(* IEC 61131-3 sources: AyCD/codesys/src/POUs, 8 files *)

(* ---- COM_UDP_RX.st ---- *)
(*
 * COM_UDP_RX - Recibe paquete UDP de Simulink (puerto 25000).
 * Deserializa T_UDP_TX_FROM_SIM (31 LREAL = 248 bytes).
 * Usa SysSocket.library (incluida en CODESYS estándar).
 *
 * Ejecutar en Task_RX cada 20 ms.
 *)
FUNCTION_BLOCK COM_UDP_RX
VAR_INPUT
    xEnable    : BOOL;
END_VAR
VAR_OUTPUT
    xConnected : BOOL;
    udiCount   : UDINT;
END_VAR
VAR
    xInit       : BOOL := FALSE;
    hSocket     : RTS_IEC_HANDLE;
    sAddr       : SOCKADDRESS;
    udiRecv     : UDINT;
    diRes       : DINT;
    abyBuffer   : ARRAY[0..255] OF BYTE;
END_VAR

(* ---- Inicialización del socket (una vez) ---- *)
IF NOT xInit AND xEnable THEN
    hSocket := SysSockCreate(SOCKET_AF_INET, SOCKET_STREAM_UDP, SOCKET_IPPROTO_UDP, ADR(diRes));
    IF diRes = 0 THEN
        // Modo no bloqueante para que Task_RX no se quede esperando
        SysSockIoctl(hSocket, SOCKET_FIONBIO, ADR(1));
        // Bind a localhost:25000
        sAddr.sin_family := SOCKET_AF_INET;
        sAddr.sin_port := SysSockHtons(GVL_PARAMS.UDP_PORT_RX);
        SysSockInetAddr('0.0.0.0', ADR(sAddr.sin_addr));
        diRes := SysSockBind(hSocket, ADR(sAddr), SIZEOF(sAddr));
        IF diRes = 0 THEN
            xInit := TRUE;
            xConnected := TRUE;
            GVL_COMMS.udp_rx_socket := SysSockHandleToDInt(hSocket);
        ELSE
            GVL_COMMS.udp_rx_err := diRes;
            SysSockClose(hSocket);
        END_IF
    ELSE
        GVL_COMMS.udp_rx_err := diRes;
    END_IF
END_IF

(* ---- Recepción no bloqueante ---- *)
IF xInit AND xEnable THEN
    udiRecv := 0;
    diRes := SysSockRecv(hSocket, ADR(abyBuffer), SIZEOF(abyBuffer), 0, ADR(udiRecv));
    IF diRes = 0 AND udiRecv = GVL_PARAMS.UDP_RX_SIZE THEN
        // Copia directa al struct (little-endian, x64)
        SysMemCpy(ADR(GVL_COMMS.udp_from_sim), ADR(abyBuffer), GVL_PARAMS.UDP_RX_SIZE);
        GVL_COMMS.udp_rx_ok := TRUE;
        GVL_COMMS.udp_rx_count := GVL_COMMS.udp_rx_count + 1;
        udiCount := GVL_COMMS.udp_rx_count;
    ELSIF diRes <> 0 AND diRes <> SOCKET_EAGAIN THEN
        GVL_COMMS.udp_rx_err := diRes;
        GVL_COMMS.udp_rx_ok := FALSE;
    END_IF
END_IF

(* ---- COM_UDP_TX.st ---- *)
(*
 * COM_UDP_TX - Envía paquete UDP a Simulink (puerto 25001).
 * Serializa T_UDP_RX_TO_SIM (53 LREAL = 424 bytes) desde GVL_COMMS.udp_to_sim.
 * Usa SysSocket.library.
 *
 * Ejecutar en Task_TX cada 20 ms (después de Task_Supervisor).
 *)
FUNCTION_BLOCK COM_UDP_TX
VAR_INPUT
    xEnable    : BOOL;
END_VAR
VAR_OUTPUT
    xConnected : BOOL;
    udiCount   : UDINT;
END_VAR
VAR
    xInit       : BOOL := FALSE;
    hSocket     : RTS_IEC_HANDLE;
    sAddrDst    : SOCKADDRESS;
    diRes       : DINT;
    udiSent     : UDINT;
    abyBuffer   : ARRAY[0..511] OF BYTE;
END_VAR

(* ---- Inicialización del socket (una vez) ---- *)
IF NOT xInit AND xEnable THEN
    hSocket := SysSockCreate(SOCKET_AF_INET, SOCKET_STREAM_UDP, SOCKET_IPPROTO_UDP, ADR(diRes));
    IF diRes = 0 THEN
        // Destino: Simulink en 127.0.0.1:25001
        sAddrDst.sin_family := SOCKET_AF_INET;
        sAddrDst.sin_port := SysSockHtons(GVL_PARAMS.UDP_PORT_TX);
        SysSockInetAddr(GVL_PARAMS.UDP_REMOTE_IP, ADR(sAddrDst.sin_addr));
        xInit := TRUE;
        xConnected := TRUE;
        GVL_COMMS.udp_tx_socket := SysSockHandleToDInt(hSocket);
    ELSE
        GVL_COMMS.udp_tx_err := diRes;
    END_IF
END_IF

(* ---- Envío cada ciclo ---- *)
IF xInit AND xEnable THEN
    // Copia struct -> buffer
    SysMemCpy(ADR(abyBuffer), ADR(GVL_COMMS.udp_to_sim), GVL_PARAMS.UDP_TX_SIZE);
    udiSent := 0;
    diRes := SysSockSendTo(hSocket, ADR(abyBuffer), GVL_PARAMS.UDP_TX_SIZE, 0,
                            ADR(sAddrDst), SIZEOF(sAddrDst), ADR(udiSent));
    IF diRes = 0 AND udiSent = GVL_PARAMS.UDP_TX_SIZE THEN
        GVL_COMMS.udp_tx_ok := TRUE;
        GVL_COMMS.udp_tx_count := GVL_COMMS.udp_tx_count + 1;
        udiCount := GVL_COMMS.udp_tx_count;
    ELSE
        GVL_COMMS.udp_tx_err := diRes;
        GVL_COMMS.udp_tx_ok := FALSE;
    END_IF
END_IF

(* ---- CONTROL_SEGURIDAD.st ---- *)
(*
 * CONTROL_SEGURIDAD (Nivel 0)
 * Capa de seguridad: watchdog, límites, emergencia, control de frenos.
 * Ejecutar en Task_Seguridad cada 20 ms.
 *
 * STUB INICIAL: estructura básica. La lógica completa de transiciones
 * debe replicar el chart Stateflow `planta/Nivel 0` de simulink/planta.slx
 *)
FUNCTION_BLOCK CONTROL_SEGURIDAD
VAR_INPUT
    // Recibidas vía COM_UDP_RX (desde GVL_COMMS.udp_from_sim)
    BTN_Emerg          : BOOL;
    BTN_Reset          : BOOL;
    FCE_der            : BOOL;
    FCE_inf            : BOOL;
    FCE_izq            : BOOL;
    FCE_sup            : BOOL;
    vh_obs             : LREAL;
    vt_obs             : LREAL;
    m_container        : LREAL;
    recup_ok           : BOOL;
    heartbeat_L1       : INT;       // pulso desde L1
END_VAR
VAR_OUTPUT
    BRK_hE_N0          : INT;       // 1 = liberado, 0 = frenado
    BRK_t_N0           : INT;
    FALLA_MAN          : BOOL;
    FALLA_WD           : BOOL;
    FALLA_IZAJE_SV     : BOOL;
    FALLA_IZAJE_INF    : BOOL;
    FALLA_IZAJE_SUP    : BOOL;
    FALLA_CARRO_DER    : BOOL;
    FALLA_CARRO_IZQ    : BOOL;
    FALLA_CARRO_SV     : BOOL;
    vh_lim             : LREAL;     // velocidad izaje límite dinámica
END_VAR
VAR
    estado             : (SISTEMA_OK, EMERG_MANUAL, EMERG_CARRO, EMERG_IZAJE,
                          EMERG_WD, MODO_RECUPERACION) := SISTEMA_OK;
    wd_state           : (WD_DOWN, WD_UP, WD_FALLO) := WD_DOWN;
    wd_counter         : DINT := 0;
    heartbeat_prev     : INT := -1;
    rTemp              : LREAL;
END_VAR

(* ============================================================
 * 1. WATCHDOG - detecta pérdida de heartbeat desde L1
 * ============================================================ *)
IF heartbeat_L1 <> heartbeat_prev THEN
    wd_state := WD_UP;
    wd_counter := 0;
    heartbeat_prev := heartbeat_L1;
ELSE
    wd_counter := wd_counter + 1;
    IF wd_counter >= GVL_PARAMS.counter_limit THEN
        wd_state := WD_FALLO;
    END_IF
END_IF

(* ============================================================
 * 2. ENVOLVENTE DE VELOCIDAD - vh_lim según masa container
 * ============================================================ *)
rTemp := GVL_PARAMS.P_nom / ((m_container + GVL_PARAMS.Ms) * GVL_PARAMS.g);
vh_lim := MIN(GVL_PARAMS.vh_max, MAX(GVL_PARAMS.vh_nom, rTemp));

(* ============================================================
 * 3. MAQUINA DE ESTADOS PRINCIPAL
 * TODO: replicar transiciones exactas del chart Stateflow.
 * Por ahora: estructura mínima funcional.
 * ============================================================ *)
CASE estado OF
    SISTEMA_OK:
        BRK_hE_N0 := 1;
        BRK_t_N0  := 1;
        FALLA_MAN := FALSE;
        FALLA_WD  := FALSE;

        IF BTN_Emerg THEN
            estado := EMERG_MANUAL;
        ELSIF wd_state = WD_FALLO THEN
            estado := EMERG_WD;
        ELSIF FCE_der OR FCE_izq THEN
            estado := EMERG_CARRO;
        ELSIF FCE_sup OR FCE_inf OR (ABS(vh_obs) > 1.15 * vh_lim) THEN
            estado := EMERG_IZAJE;
        END_IF

    EMERG_MANUAL:
        BRK_hE_N0 := 0;
        BRK_t_N0  := 0;
        FALLA_MAN := TRUE;
        IF NOT BTN_Emerg AND BTN_Reset THEN
            estado := MODO_RECUPERACION;
        END_IF

    EMERG_CARRO:
        BRK_hE_N0 := 1;        // izaje libre
        BRK_t_N0  := 0;        // carro frenado
        FALLA_CARRO_DER := FCE_der;
        FALLA_CARRO_IZQ := FCE_izq;
        IF BTN_Reset THEN
            estado := MODO_RECUPERACION;
        END_IF

    EMERG_IZAJE:
        BRK_hE_N0 := 0;
        BRK_t_N0  := 1;
        FALLA_IZAJE_INF := FCE_inf;
        FALLA_IZAJE_SUP := FCE_sup;
        FALLA_IZAJE_SV  := ABS(vh_obs) > 1.15 * vh_lim;
        IF BTN_Reset THEN
            estado := MODO_RECUPERACION;
        END_IF

    EMERG_WD:
        BRK_hE_N0 := 0;
        BRK_t_N0  := 0;
        FALLA_WD  := TRUE;
        IF wd_state <> WD_FALLO AND BTN_Reset THEN
            estado := MODO_RECUPERACION;
        END_IF

    MODO_RECUPERACION:
        BRK_hE_N0 := 0;
        BRK_t_N0  := 0;
        IF recup_ok THEN
            FALLA_MAN := FALSE;
            FALLA_WD  := FALSE;
            FALLA_IZAJE_INF := FALSE;
            FALLA_IZAJE_SUP := FALSE;
            FALLA_IZAJE_SV  := FALSE;
            FALLA_CARRO_DER := FALSE;
            FALLA_CARRO_IZQ := FALSE;
            FALLA_CARRO_SV  := FALSE;
            estado := SISTEMA_OK;
        END_IF
END_CASE

(* ============================================================
 * 4. Publicar a GVL_PROCESS para que L1 lea
 * ============================================================ *)
GVL_PROCESS.FALLA_GLOBAL := FALLA_MAN OR FALLA_WD OR FALLA_IZAJE_SV
                          OR FALLA_IZAJE_INF OR FALLA_IZAJE_SUP
                          OR FALLA_CARRO_DER OR FALLA_CARRO_IZQ OR FALLA_CARRO_SV;
GVL_PROCESS.FALLA_MAN_L0       := FALLA_MAN;
GVL_PROCESS.FALLA_WD_L0        := FALLA_WD;
GVL_PROCESS.FALLA_SV_L0        := FALLA_IZAJE_SV;
GVL_PROCESS.FALLA_CARRO_DER_L0 := FALLA_CARRO_DER;
GVL_PROCESS.FALLA_CARRO_IZQ_L0 := FALLA_CARRO_IZQ;
GVL_PROCESS.FALLA_CARRO_SV_L0  := FALLA_CARRO_SV;
GVL_PROCESS.FALLA_IZAJE_INF_L0 := FALLA_IZAJE_INF;
GVL_PROCESS.FALLA_IZAJE_SUP_L0 := FALLA_IZAJE_SUP;
GVL_PROCESS.FALLA_IZAJE_SV_L0  := FALLA_IZAJE_SV;
GVL_PROCESS.RECUPERAR_L0       := (estado = MODO_RECUPERACION);
GVL_PROCESS.vh_lim_L0          := vh_lim;
GVL_PROCESS.BRK_h_N0           := BRK_hE_N0;
GVL_PROCESS.BRK_t_N0           := BRK_t_N0;

(* ---- CONTROL_SUPERVISOR.st ---- *)
(*
 * CONTROL_SUPERVISOR (Nivel 1)
 * Capa de supervisión: máquina principal manual/auto/error, twistlocks,
 * generación de heartbeat, suavizado cinemático, selección de trayectoria.
 * Ejecutar en Task_Supervisor cada 20 ms.
 *
 * STUB INICIAL: estructura básica. La lógica completa debe replicar
 * el chart Stateflow `planta/Nivel 1` de simulink/planta.slx
 *)
FUNCTION_BLOCK CONTROL_SUPERVISOR
VAR_INPUT
    // Recibidas vía COM_UDP_RX (desde GVL_COMMS.udp_from_sim)
    BTN_ON_OFF         : BOOL;
    BTN_TLK            : BOOL;
    BTN_Auto           : BOOL;
    BTN_Reset          : BOOL;
    Joy_XY             : ARRAY[1..2] OF LREAL;
    theta_l            : LREAL;
    theta_l_dot        : LREAL;
    vh_obs             : LREAL;
    vt_obs             : LREAL;
    Fhw                : LREAL;
    yh_enc             : LREAL;
    xt_enc             : LREAL;
    FC_der             : BOOL;
    FC_inf             : BOOL;
    FC_izq             : BOOL;
    FC_sup             : BOOL;
    T_hm               : LREAL;
    T_tm               : LREAL;
    // De L0 (vía GVL_PROCESS)
    FALLA_GLOBAL       : BOOL;
    RECUPERAR_L0       : BOOL;
END_VAR
VAR_OUTPUT
    BRK_h_N1           : INT;
    BRK_t_N1           : INT;
    TLK_OUT            : INT;
    yc0_vec_OUT        : ARRAY[1..33] OF LREAL;
    i_sel_OUT          : LREAL;
    vx_suave           : LREAL;
    vy_suave           : LREAL;
    recuperacion_OUT   : BOOL;
    modo_muerto        : BOOL;
    heartbeat_OUT      : INT;
    m_container_OUT    : LREAL;
END_VAR
VAR
    estado             : (STAND_BY, MANUAL, AUTO, PASO_STAND_BY,
                          ERROR_GENERICO, RECUPERACION) := STAND_BY;
    sub_auto           : (AUTO_INIT, SEL_INDICE_INI, SEL_INDICE_FIN,
                          SEL_TRAYECTORIA, MOV_CURVO, MOV_SEGURO,
                          MANUAL_SIMPLE) := AUTO_INIT;
    twistlock          : (TLK_VACIO, TLK_CERRANDO, TLK_CARGADO,
                          TLK_ABRIENDO) := TLK_VACIO;
    heartbeat_int      : INT := 0;
    i_origen           : INT := 0;
    i_destino          : INT := 0;
    i_sel              : INT := 1;
    cont_valido        : BOOL := FALSE;
    tlk_cerrado        : BOOL := FALSE;
    rAcc               : LREAL := 0.0;
    yc0_vec_initialized: BOOL := FALSE;
END_VAR

(* ============================================================
 * 1. INIT - cargar perfil inicial (una vez)
 * ============================================================ *)
IF NOT yc0_vec_initialized THEN
    (* Perfil inicial de containers (espejo h_vec_inicial * Hc en init_plant_parameters.m).
       Valores escalados por Hc=2.59. Editar si difieren los del chart Stateflow real. *)
    yc0_vec_OUT[1]  := 0.0;
    yc0_vec_OUT[2]  := 0.0;
    yc0_vec_OUT[3]  := GVL_PARAMS.Hc;
    yc0_vec_OUT[4]  := 0.0;
    yc0_vec_OUT[5]  := 0.0;
    yc0_vec_OUT[6]  := GVL_PARAMS.Hc;
    yc0_vec_OUT[7]  := 0.0;
    yc0_vec_OUT[8]  := 0.0;
    yc0_vec_OUT[9]  := 0.0;
    yc0_vec_OUT[10] := 0.0;
    yc0_vec_OUT[11] := 0.0;
    yc0_vec_OUT[12] := 0.0;
    yc0_vec_OUT[13] := GVL_PARAMS.alt_borde * GVL_PARAMS.Hc;
    yc0_vec_OUT[14] := 3.0 * GVL_PARAMS.Hc;
    yc0_vec_OUT[15] := 5.0 * GVL_PARAMS.Hc;
    yc0_vec_OUT[16] := 6.0 * GVL_PARAMS.Hc;
    yc0_vec_OUT[17] := 3.0 * GVL_PARAMS.Hc;
    yc0_vec_OUT[18] := 5.0 * GVL_PARAMS.Hc;
    yc0_vec_OUT[19] := 6.0 * GVL_PARAMS.Hc;
    yc0_vec_OUT[20] := 6.0 * GVL_PARAMS.Hc;
    yc0_vec_OUT[21] := 4.0 * GVL_PARAMS.Hc;
    yc0_vec_OUT[22] := 1.0 * GVL_PARAMS.Hc;
    yc0_vec_OUT[23] := 1.0 * GVL_PARAMS.Hc;
    yc0_vec_OUT[24] := -4.0 * GVL_PARAMS.Hc;
    yc0_vec_OUT[25] := -5.0 * GVL_PARAMS.Hc;
    yc0_vec_OUT[26] := -2.0 * GVL_PARAMS.Hc;
    yc0_vec_OUT[27] := -1.0 * GVL_PARAMS.Hc;
    yc0_vec_OUT[28] := 2.0 * GVL_PARAMS.Hc;
    yc0_vec_OUT[29] := 6.0 * GVL_PARAMS.Hc;
    yc0_vec_OUT[30] := 4.0 * GVL_PARAMS.Hc;
    yc0_vec_OUT[31] := 2.0 * GVL_PARAMS.Hc;
    yc0_vec_OUT[32] := 5.0 * GVL_PARAMS.Hc;
    yc0_vec_OUT[33] := GVL_PARAMS.alt_borde * GVL_PARAMS.Hc;
    yc0_vec_initialized := TRUE;
END_IF

(* ============================================================
 * 2. HEARTBEAT - toggle por ciclo para el watchdog de L0
 * ============================================================ *)
IF heartbeat_int = 0 THEN
    heartbeat_int := 1;
ELSE
    heartbeat_int := 0;
END_IF
heartbeat_OUT := heartbeat_int;
GVL_PROCESS.heartbeat_L1 := heartbeat_int;

(* ============================================================
 * 3. ESTIMACION DE MASA - cuando twistlock cerrado y carga colgando
 * TODO: replicar lógica del chart Stateflow
 * ============================================================ *)
IF tlk_cerrado THEN
    m_container_OUT := MAX(0.0, ABS(Fhw) / GVL_PARAMS.g - GVL_PARAMS.Ms);
ELSE
    m_container_OUT := 0.0;
END_IF
GVL_PROCESS.m_container_L1 := m_container_OUT;

(* ============================================================
 * 4. MAQUINA TWISTLOCKS (paralela a la principal)
 * ============================================================ *)
CASE twistlock OF
    TLK_VACIO:
        TLK_OUT := 0;
        IF BTN_TLK AND ABS(Fhw) > 100.0 THEN
            twistlock := TLK_CERRANDO;
        END_IF
    TLK_CERRANDO:
        TLK_OUT := 1;
        tlk_cerrado := TRUE;
        twistlock := TLK_CARGADO;
    TLK_CARGADO:
        TLK_OUT := 1;
        IF BTN_TLK AND ABS(Fhw) < 100.0 THEN
            twistlock := TLK_ABRIENDO;
        END_IF
    TLK_ABRIENDO:
        TLK_OUT := 0;
        tlk_cerrado := FALSE;
        twistlock := TLK_VACIO;
END_CASE

(* ============================================================
 * 5. MAQUINA PRINCIPAL
 * STUB - replicar transiciones exactas del chart Stateflow
 * ============================================================ *)
CASE estado OF
    STAND_BY:
        BRK_h_N1 := 0;
        BRK_t_N1 := 0;
        vx_suave := 0.0;
        vy_suave := 0.0;
        modo_muerto := TRUE;
        IF FALLA_GLOBAL THEN
            estado := ERROR_GENERICO;
        ELSIF BTN_ON_OFF AND NOT BTN_Auto THEN
            estado := MANUAL;
        ELSIF BTN_Auto THEN
            estado := AUTO;
            sub_auto := AUTO_INIT;
        END_IF

    MANUAL:
        BRK_h_N1 := 1;
        BRK_t_N1 := 1;
        modo_muerto := FALSE;
        // Aplicar zona muerta al joystick
        IF ABS(Joy_XY[1]) > GVL_PARAMS.dead_zone THEN
            vx_suave := Joy_XY[1] * GVL_PARAMS.vt_max;
        ELSE
            vx_suave := 0.0;
        END_IF
        IF ABS(Joy_XY[2]) > GVL_PARAMS.dead_zone THEN
            vy_suave := Joy_XY[2] * GVL_PARAMS.vh_max;
        ELSE
            vy_suave := 0.0;
        END_IF
        IF FALLA_GLOBAL THEN
            estado := ERROR_GENERICO;
        ELSIF NOT BTN_ON_OFF THEN
            estado := STAND_BY;
        END_IF

    AUTO:
        BRK_h_N1 := 1;
        BRK_t_N1 := 1;
        modo_muerto := FALSE;
        // Sub-máquina (TODO: completar transiciones reales)
        CASE sub_auto OF
            AUTO_INIT:
                sub_auto := SEL_INDICE_INI;
            SEL_INDICE_INI:
                IF ABS(Joy_XY[1]) > GVL_PARAMS.dead_zone THEN
                    // ajustar índice según signo del joystick
                    ;
                END_IF
                IF BTN_TLK THEN
                    i_origen := i_sel;
                    sub_auto := SEL_INDICE_FIN;
                END_IF
            SEL_INDICE_FIN:
                IF BTN_TLK THEN
                    i_destino := i_sel;
                    sub_auto := SEL_TRAYECTORIA;
                END_IF
            SEL_TRAYECTORIA:
                sub_auto := MOV_CURVO;
            MOV_CURVO:
                // mover hasta i_destino
                ;
            MOV_SEGURO:
                ;
            MANUAL_SIMPLE:
                ;
        END_CASE
        IF FALLA_GLOBAL THEN
            estado := ERROR_GENERICO;
        ELSIF NOT BTN_Auto THEN
            estado := PASO_STAND_BY;
        END_IF
        i_sel_OUT := DINT_TO_LREAL(i_sel);

    PASO_STAND_BY:
        vx_suave := 0.0;
        vy_suave := 0.0;
        IF ABS(vh_obs) < 0.01 AND ABS(vt_obs) < 0.01 THEN
            estado := STAND_BY;
        END_IF

    ERROR_GENERICO:
        BRK_h_N1 := 0;
        BRK_t_N1 := 0;
        vx_suave := 0.0;
        vy_suave := 0.0;
        modo_muerto := TRUE;
        IF RECUPERAR_L0 THEN
            estado := RECUPERACION;
        END_IF

    RECUPERACION:
        // Mover a posición segura (TODO: lógica completa)
        recuperacion_OUT := TRUE;
        IF NOT FALLA_GLOBAL THEN
            recuperacion_OUT := FALSE;
            estado := STAND_BY;
        END_IF
END_CASE

(* ============================================================
 * 6. Publicar a GVL_PROCESS y GVL_COMMS.udp_to_sim
 * ============================================================ *)
GVL_PROCESS.BRK_h_N1         := BRK_h_N1;
GVL_PROCESS.BRK_t_N1         := BRK_t_N1;
GVL_PROCESS.TLK_OUT          := TLK_OUT;
GVL_PROCESS.vx_suave         := vx_suave;
GVL_PROCESS.vy_suave         := vy_suave;
GVL_PROCESS.i_sel_OUT        := i_sel;
GVL_PROCESS.recuperacion_OUT := recuperacion_OUT;
GVL_PROCESS.modo_muerto_L1   := modo_muerto;
GVL_PROCESS.yc0_vec_OUT      := yc0_vec_OUT;

(* ---- PRG_RX.st ---- *)
(*
 * PRG_RX - Programa llamado por Task_RX (20 ms).
 * Recibe UDP de Simulink y mapea los campos al GVL_COMMS.udp_from_sim.
 *)
PROGRAM PRG_RX
VAR
    fbUdpRx : COM_UDP_RX;
END_VAR

fbUdpRx(xEnable := TRUE);

(* ---- PRG_SEGURIDAD.st ---- *)
(*
 * PRG_SEGURIDAD - Programa llamado por Task_Seguridad (20 ms).
 * Desempaqueta entradas y ejecuta CONTROL_SEGURIDAD (L0).
 *)
PROGRAM PRG_SEGURIDAD
VAR
    fbSeguridad : CONTROL_SEGURIDAD;
END_VAR

fbSeguridad(
    BTN_Emerg     := GVL_COMMS.udp_from_sim.BTN_Emerg > 0.5,
    BTN_Reset     := GVL_COMMS.udp_from_sim.BTN_Reset > 0.5,
    FCE_der       := GVL_COMMS.udp_from_sim.FCE_der > 0.5,
    FCE_inf       := GVL_COMMS.udp_from_sim.FCE_inf > 0.5,
    FCE_izq       := GVL_COMMS.udp_from_sim.FCE_izq > 0.5,
    FCE_sup       := GVL_COMMS.udp_from_sim.FCE_sup > 0.5,
    vh_obs        := GVL_COMMS.udp_from_sim.vh_obs,
    vt_obs        := GVL_COMMS.udp_from_sim.vt_obs,
    m_container   := GVL_PROCESS.m_container_L1,
    recup_ok      := GVL_COMMS.udp_from_sim.recup_ok > 0.5,
    heartbeat_L1  := GVL_PROCESS.heartbeat_L1
);

(* ---- PRG_SUPERVISOR.st ---- *)
(*
 * PRG_SUPERVISOR - Programa llamado por Task_Supervisor (20 ms).
 * Desempaqueta entradas y ejecuta CONTROL_SUPERVISOR (L1).
 *)
PROGRAM PRG_SUPERVISOR
VAR
    fbSupervisor : CONTROL_SUPERVISOR;
END_VAR

fbSupervisor(
    BTN_ON_OFF    := GVL_COMMS.udp_from_sim.BTN_ON_OFF > 0.5,
    BTN_TLK       := GVL_COMMS.udp_from_sim.BTN_TLK > 0.5,
    BTN_Auto      := GVL_COMMS.udp_from_sim.BTN_Auto > 0.5,
    BTN_Reset     := GVL_COMMS.udp_from_sim.BTN_Reset > 0.5,
    Joy_XY        := GVL_COMMS.udp_from_sim.Joy_XY,
    theta_l       := GVL_COMMS.udp_from_sim.theta_l,
    theta_l_dot   := GVL_COMMS.udp_from_sim.theta_l_dot,
    vh_obs        := GVL_COMMS.udp_from_sim.vh_obs,
    vt_obs        := GVL_COMMS.udp_from_sim.vt_obs,
    Fhw           := GVL_COMMS.udp_from_sim.Fhw,
    yh_enc        := GVL_COMMS.udp_from_sim.yh_enc,
    xt_enc        := GVL_COMMS.udp_from_sim.xt_enc,
    FC_der        := GVL_COMMS.udp_from_sim.FC_der > 0.5,
    FC_inf        := GVL_COMMS.udp_from_sim.FC_inf > 0.5,
    FC_izq        := GVL_COMMS.udp_from_sim.FC_izq > 0.5,
    FC_sup        := GVL_COMMS.udp_from_sim.FC_sup > 0.5,
    T_hm          := GVL_COMMS.udp_from_sim.T_hm,
    T_tm          := GVL_COMMS.udp_from_sim.T_tm,
    FALLA_GLOBAL  := GVL_PROCESS.FALLA_GLOBAL,
    RECUPERAR_L0  := GVL_PROCESS.RECUPERAR_L0
);

(* ---- PRG_TX.st ---- *)
(*
 * PRG_TX - Programa llamado por Task_TX (20 ms).
 * Empaqueta señales del PLC en GVL_COMMS.udp_to_sim y las envía.
 *)
PROGRAM PRG_TX
VAR
    fbUdpTx : COM_UDP_TX;
END_VAR

(* Empaquetar valores actuales del PLC en el struct de salida *)
GVL_COMMS.udp_to_sim.BRK_h_N1        := INT_TO_LREAL(GVL_PROCESS.BRK_h_N1);
GVL_COMMS.udp_to_sim.BRK_t_N1        := INT_TO_LREAL(GVL_PROCESS.BRK_t_N1);
GVL_COMMS.udp_to_sim.TLK             := INT_TO_LREAL(GVL_PROCESS.TLK_OUT);
GVL_COMMS.udp_to_sim.yc0_vec         := GVL_PROCESS.yc0_vec_OUT;
GVL_COMMS.udp_to_sim.i_sel           := INT_TO_LREAL(GVL_PROCESS.i_sel_OUT);
GVL_COMMS.udp_to_sim.vx_suave        := GVL_PROCESS.vx_suave;
GVL_COMMS.udp_to_sim.vy_suave        := GVL_PROCESS.vy_suave;
GVL_COMMS.udp_to_sim.recuperacion    := BOOL_TO_LREAL(GVL_PROCESS.recuperacion_OUT);
GVL_COMMS.udp_to_sim.modo_muerto     := BOOL_TO_LREAL(GVL_PROCESS.modo_muerto_L1);
GVL_COMMS.udp_to_sim.heartbeat       := INT_TO_LREAL(GVL_PROCESS.heartbeat_L1);
GVL_COMMS.udp_to_sim.m_container     := GVL_PROCESS.m_container_L1;
GVL_COMMS.udp_to_sim.BRK_hE_N0       := INT_TO_LREAL(GVL_PROCESS.BRK_h_N0);
GVL_COMMS.udp_to_sim.BRK_t_N0        := INT_TO_LREAL(GVL_PROCESS.BRK_t_N0);
GVL_COMMS.udp_to_sim.FALLA_IZAJE_SV  := BOOL_TO_LREAL(GVL_PROCESS.FALLA_IZAJE_SV_L0);
GVL_COMMS.udp_to_sim.FALLA_MAN       := BOOL_TO_LREAL(GVL_PROCESS.FALLA_MAN_L0);
GVL_COMMS.udp_to_sim.FALLA_WD        := BOOL_TO_LREAL(GVL_PROCESS.FALLA_WD_L0);
GVL_COMMS.udp_to_sim.FALLA_CARRO_DER := BOOL_TO_LREAL(GVL_PROCESS.FALLA_CARRO_DER_L0);
GVL_COMMS.udp_to_sim.FALLA_CARRO_IZQ := BOOL_TO_LREAL(GVL_PROCESS.FALLA_CARRO_IZQ_L0);
GVL_COMMS.udp_to_sim.FALLA_IZAJE_INF := BOOL_TO_LREAL(GVL_PROCESS.FALLA_IZAJE_INF_L0);
GVL_COMMS.udp_to_sim.FALLA_IZAJE_SUP := BOOL_TO_LREAL(GVL_PROCESS.FALLA_IZAJE_SUP_L0);
GVL_COMMS.udp_to_sim.FALLA_CARRO_SV  := BOOL_TO_LREAL(GVL_PROCESS.FALLA_CARRO_SV_L0);

fbUdpTx(xEnable := TRUE);
